Fanuc KAREL source: kb00160.KL

-- PROVISIONAL review KL for V1013-1; original PC SHA256 eb6a5129c7e0160ceec51766e47608f6387f982a23d01cf5865fa628b4b626bb
-- Incomplete behavior may be omitted. Consult companion uncertainty JSON. Do not deploy.
PROGRAM KB00160
%NOLOCKGROUP
BEGIN
  -- UNRESOLVED_PC offsets 5-12; opcodes 9D,23
  -- UNRESOLVED_PC offsets 17-24; opcodes 9D,23
  -- UNRESOLVED_PC offsets 29-36; opcodes 9D,23
  -- UNRESOLVED_PC offsets 41-69; opcodes 27,22,22,22,22,31
  -- UNRESOLVED_PC offsets 74-78; opcodes 7F
END KB00160
